RoboDK station: RobodkBasico-2.rdk

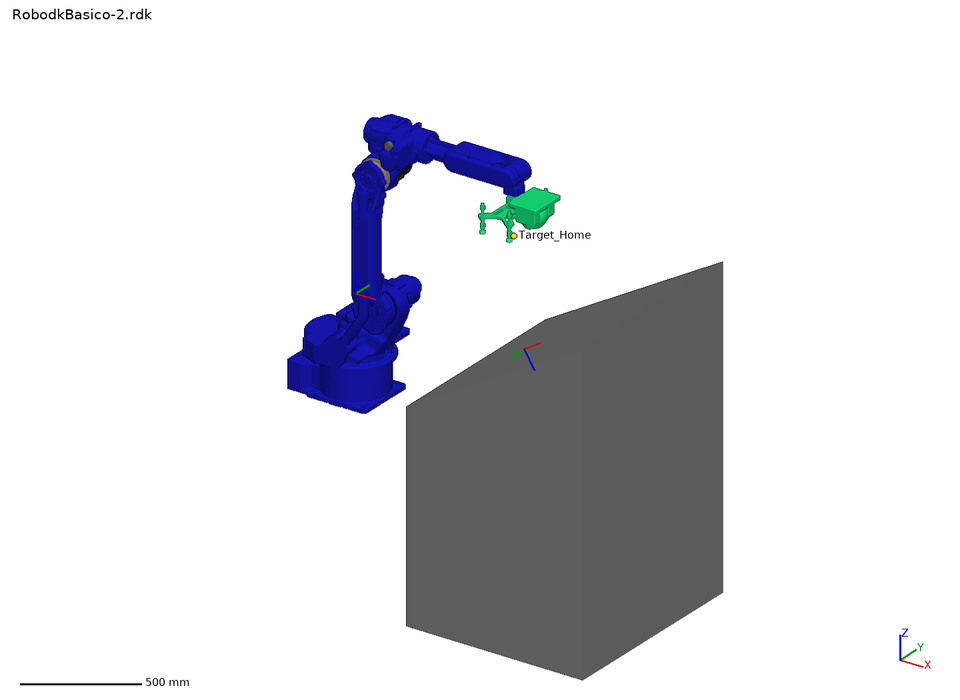
[picture v0: the station drawn from its stored meshes, robots at their saved joint values, targets as dots, program paths as lines]
Station Robodk (2) (saved by RoboDK 6.1.1). Poses are relative to the parent item; angles as X-Y-Z fixed-axis rotations.
  - frame Motoman MH6 Base at (0, 0, 450) mm
    - robot Motoman MH6: 6 axes, payload 6 kg, reach 1422 mm, repeatability 0.08 mm, weight 130 kg
        modified DH rows (alpha deg, a mm, theta deg, d mm): 0, 0, 0, 450; -90, 152, -90, 0; 0, 614, 0, 0; -90, 155, 0, 640; 90, 0, 90, 0; -90, 0, 0, 95
        base shift (0, 0, -450) mm
        joint limits [-170, -90, -175, -180, -45, -360] to [170, 155, 250, 180, 225, 360]; home [0, 0, 0, 0, 0, 0]; saved at [0, 0, 0, 0, 0, 0]
      - tool Ventosas, TCP at (0, 0, 190) mm, size 250 x 290 x 148 mm
    - frame Frame_from_Target1 at (866.5, -34.49, 3.87) mm, rotated rx -180 ry -30 rz 0 deg
      - target Target_Home (Cartesian target) at (175.55, -34.49, -453.06) mm, rotated rx 0 ry -30 rz 0 deg; joints [0, 0, 0, 0, 0, 0] of Motoman MH6
  - object CAJA2 at (1600, 500, 300) mm, rotated rx 180 ry 0 rz 0 deg, size 886.4 x 1000 x 1511.7 mm, geometry from CAJA2.stp
  - Python program RosPolar (listed below)

--- Python program RosPolar ---
from robodk.robolink import *    # API para comunicarte con RoboDK
from robodk.robomath import *    # Funciones matemáticas
import math
from matplotlib.textpath import TextPath
from matplotlib.font_manager import FontProperties

#------------------------------------------------
# 1) Conexión a RoboDK e inicialización
#------------------------------------------------
RDK = Robolink()

# Elegir un robot (si hay varios, aparece un popup)
robot = RDK.ItemUserPick("Selecciona un robot", ITEM_TYPE_ROBOT)
if not robot.Valid():
    raise Exception("No se ha seleccionado un robot válido.")

### Conectar al robot físico
##if not robot.Connect():
##    raise Exception("No se pudo conectar al robot. Verifica que esté en modo remoto y que la configuración sea correcta.")
##
### Confirmar conexión
##if not robot.ConnectedState():
##    raise Exception("El robot no está conectado correctamente. Revisa la conexión.")
##
##print("Robot conectado correctamente.")

#------------------------------------------------
# 2) Cargar el Frame (ya existente) donde quieres dibujar
#    Ajusta el nombre si tu Frame se llama diferente
#------------------------------------------------
frame_name = "Frame_from_Target1"
frame = RDK.Item(frame_name, ITEM_TYPE_FRAME)
if not frame.Valid():
    raise Exception(f'No se encontró el Frame "{frame_name}" en la estación.')

# Asignamos este frame al robot
robot.setPoseFrame(frame)
# Usamos la herramienta activa
robot.setPoseTool(robot.PoseTool())

# Ajustes de velocidad y blending
robot.setSpeed(80)   # mm/s - Ajusta según necesites
robot.setRounding(5)  # blending (radio de curvatura)

#####################################################################
# Movimiento a Home

nombre_home = "Target_Home"
T_H = RDK.Item(nombre_home, ITEM_TYPE_TARGET)
if not T_H.Valid():
    raise Exception(f'No se encontró el target "{nombre_home}" en la estación.')

def ir_a_home():
    robot.MoveJ(T_H)

ir_a_home()

#------------------------------------------------
# 3) Parámetros de la figura (rosa polar)
#------------------------------------------------
n, d = 1, 4
num_points = 720       # Cuántos puntos muestreamos (mayor = más suave)
A = 110                # Amplitud (300 mm = radio máximo)
k = n/d                # Parámetro de la rosa (pétalos). Si es impar, habrá k pétalos; si es par, 2k
theta_max = math.pi * d if (n * d) % 2 == 1 else 2 * math.pi * d
z_surface = 0          # Z=0 en el plano del frame
z_safe = 50            # Altura segura para aproximarse y salir
z_up = z_surface - z_safe

ANGULO = -90
ESPEJO_X = True
OFFSET_X = 0
OFFSET_Y = 0

_c = math.cos(math.radians(ANGULO))
_s = math.sin(math.radians(ANGULO))

def transformar(x, y):
    if ESPEJO_X:
        x = -x
    xr = x * _c - y * _s
    yr = x * _s + y * _c
    return xr + OFFSET_X, yr + OFFSET_Y

def trazo(puntos):
    puntos = [transformar(x, y) for x, y in puntos]
    x0, y0 = puntos[0]
    robot.MoveL(transl(x0, y0, z_up))
    robot.MoveL(transl(x0, y0, z_surface))
    for j, (x, y) in enumerate(puntos[1:], start=1):
        try:
            robot.MoveL(transl(x, y, z_surface))
        except Exception:
            print(f"Falla en el punto {j}: x={x:.1f}, y={y:.1f}")
            raise
    x1, y1 = puntos[-1]
    robot.MoveL(transl(x1, y1, z_up))

# Recorrido a puntos de la figura polar

rosa = []
for i in range(num_points + 1):
    theta = theta_max * i / num_points
    r = A * math.cos(k * theta)
    rosa.append((r * math.cos(theta), r * math.sin(theta)))

y_min = min(p[1] for p in rosa)

# Nombre

nombre = "Tito & Juan"
tam_fuente = 40      # mm aprox.; controla el tamaño del texto
margen = 25          # mm entre la rosa y el texto

fp = FontProperties(family="DejaVu Sans", weight="bold")
tp = TextPath((0, 0), nombre, size=tam_fuente, prop=fp)

# Contornos aplanados (las curvas Bézier quedan convertidas en segmentos)
contornos = tp.to_polygons(closed_only=False)

# Para centrar en x = 0 y ubicar el texto debajo de la rosa
ext = tp.get_extents()
dx = -(ext.x0 + ext.x1) / 2          # centrado horizontal
dy = (y_min - margen) - ext.y1       # la parte alta del texto queda bajo la rosa

texto_trazos = []
for c in contornos:
    pts = [(float(px) + dx, float(py) + dy) for px, py in c]
    if pts[0] != pts[-1]:            # cierra el contorno si no vino cerrado
        pts.append(pts[0])
    texto_trazos.append(pts)

# DIBUJO

# Aproximación sobre el inicio de la rosa (A, 0)
robot.MoveJ(transl(rosa[0][0], rosa[0][1], z_up))
trazo(rosa)

for pts in texto_trazos:
    trazo(pts)

#############################################################
# Movimiento a Home para terminar
print("Volviendo a posicion HOME")
ir_a_home()


print(f"¡Figura polar completada en el frame '{frame_name}'!")
